(* IEC 61131-3 sources: llm-plc-st-eval/data/processed_v2_primera/gpt-4o/B1/few_shot, 3 files *)

(* ---- ejec_1.st ---- *)
FUNCTION_BLOCK FB_Motor
VAR_INPUT
    btnMarcha : BOOL; (* Botón de marcha *)
    btnParo : BOOL;   (* Botón de paro *)
    btnEmerg : BOOL;  (* Botón de paro de emergencia *)
END_VAR
VAR_OUTPUT
    motorOn : BOOL;   (* Estado del motor *)
END_VAR
VAR
    motorLatch : BOOL; (* Latch para mantener el estado del motor *)
END_VAR

(* Control de arranque y paro del motor *)
IF btnEmerg THEN
    motorLatch := FALSE; (* Paro de emergencia, motor no rearranca *)
ELSIF btnParo THEN
    motorLatch := FALSE; (* Paro normal, motor se apaga *)
ELSIF btnMarcha THEN
    motorLatch := TRUE;  (* Arranque del motor, se mantiene encendido *)
END_IF

motorOn := motorLatch; (* Salida del estado del motor *)
END_FUNCTION_BLOCK

(* ---- ejec_2.st ---- *)
FUNCTION_BLOCK FB_Motor
VAR_INPUT
    btnMarcha : BOOL; (* Botón de marcha *)
    btnParo : BOOL;   (* Botón de paro *)
    btnEmerg : BOOL;  (* Botón de paro de emergencia *)
END_VAR
VAR_OUTPUT
    motorOn : BOOL;   (* Estado del motor *)
END_VAR
VAR
    motorLatch : BOOL; (* Latch para mantener el motor encendido *)
END_VAR

(* Control de arranque y paro del motor *)
IF btnEmerg THEN
    motorLatch := FALSE; (* Paro de emergencia, motor no rearranca *)
ELSIF btnParo THEN
    motorLatch := FALSE; (* Paro normal, motor se apaga *)
ELSIF btnMarcha THEN
    motorLatch := TRUE;  (* Arranque del motor *)
END_IF;

motorOn := motorLatch; (* Actualización del estado del motor *)
END_FUNCTION_BLOCK

(* ---- ejec_3.st ---- *)
FUNCTION_BLOCK FB_Motor
VAR_INPUT
    btnMarcha : BOOL; (* Botón de marcha *)
    btnParo : BOOL;   (* Botón de paro *)
    btnEmerg : BOOL;  (* Botón de paro de emergencia *)
END_VAR
VAR_OUTPUT
    motorOn : BOOL;   (* Estado del motor *)
END_VAR
VAR
    estadoEmergencia : BOOL; (* Indica si hubo un paro de emergencia *)
END_VAR

(* Si se presiona el botón de emergencia, se activa el estado de emergencia *)
IF btnEmerg THEN
    estadoEmergencia := TRUE;
END_IF

(* Si no hay estado de emergencia, el motor se enciende con el botón de marcha y se apaga con el botón de paro *)
IF NOT estadoEmergencia THEN
    IF btnMarcha THEN
        motorOn := TRUE;
    END_IF;
    IF btnParo THEN
        motorOn := FALSE;
    END_IF;
ELSE
    (* Si hay estado de emergencia, el motor se apaga y no puede rearrancar *)
    motorOn := FALSE;
END_IF;
END_FUNCTION_BLOCK
